(* IEC 61131-3 sources: codesys-framework/txt/application/ToDo/Hardware/IO/Camera/I_Camera, 9 files *)

(* ---- Connect.method.st ---- *)
METHOD Connect : BOOL
VAR_INPUT
END_VAR

(* ---- ConnectMethod.method.st ---- *)
METHOD PUBLIC ConnectMethod : BOOL
VAR_INPUT
END_VAR

(* ---- Disconnect.method.st ---- *)
METHOD Disconnect : BOOL
VAR_INPUT
END_VAR

(* ---- GetResult.method.st ---- *)
METHOD GetResult : STRING(255)
VAR_INPUT
END_VAR

(* ---- Initialize.method.st ---- *)
METHOD Initialize
VAR_INPUT
END_VAR

(* ---- Reset.method.st ---- *)
METHOD Reset
VAR_INPUT
END_VAR

(* ---- ResetResult.method.st ---- *)
METHOD ResetResult
VAR_INPUT
END_VAR

(* ---- SetJob.method.st ---- *)
METHOD SetJob : BOOL
VAR_INPUT
	id 		: UINT;
END_VAR

(* ---- TakePicture.method.st ---- *)
METHOD TakePicture : BOOL
VAR_INPUT
	pictureId		: STRING;
END_VAR
